   #FRK_Route_DeclarationCell := FALSE;
   IF NOT "FRK_PathOwned"(OwnerPath := #Module.Status.Name, TargetPath := #Request.TargetPath) THEN
       RETURN;
   END_IF;
   IF #Request.TargetPath = STRING_TO_WSTRING(#Module.Status.Name) THEN
       FOR #Index := 1 TO 16 DO
           #Module.ManConditions[#Index].Used := FALSE;
       END_FOR;
       "FRK_ManualApply"(Core := #Module.Core,
                         Status := #Module.Status,
                         Request := #Request,
                         Commands := #Module.Catalog,
                         Count := #Module.CatalogCount,
                         Conditions := #Module.ManConditions,
                         Report := #Report,
                         Execute := #Module.Execute,
                         Command := #Module.Command,
                         ManualOwned := #Module.ManualOwned);
       #FRK_Route_DeclarationCell := TRUE;
       RETURN;
   END_IF;
   #RouteMatched := "FRK_Route_DeclarationCylinder"(Module := #Module.Clamp, Hal := #Hal.Clamp, Request := #Request, Report := #Report);
   #FRK_Route_DeclarationCell := #FRK_Route_DeclarationCell OR #RouteMatched;
   #RouteMatched := "FRK_Route_DeclarationCylinder"(Module := #Module.Gate, Hal := #Hal.Gate, Request := #Request, Report := #Report);
   #FRK_Route_DeclarationCell := #FRK_Route_DeclarationCell OR #RouteMatched;
END_FUNCTION

FUNCTION "FRK_Route_DeclarationCylinder" : Bool   // FC130, SCL
{ S7_Optimized_Access := 'TRUE' }
VERSION : 0.1
// stored: AutoNumber true, IsIECCheckEnabled false, SetENOAutomatically false, UDAEnableTagReadback false
   VAR_INPUT
      Request : "ST_HmiRequest";
   END_VAR
   VAR_IN_OUT
      Module : "FB_DeclarationCylinder";
      Hal : "ST_DeclarationLeafHal";
      Report : "ST_ReleaseReport";
   END_VAR
   VAR_TEMP
      RouteMatched : Bool;
      Index : Int;
   END_VAR
BEGIN

   #FRK_Route_DeclarationCylinder := FALSE;
   IF NOT "FRK_PathOwned"(OwnerPath := #Module.Status.Name, TargetPath := #Request.TargetPath) THEN
       RETURN;
   END_IF;
   IF #Request.TargetPath = STRING_TO_WSTRING(#Module.Status.Name) THEN
       FOR #Index := 1 TO 16 DO
           #Module.ManConditions[#Index].Used := FALSE;
       END_FOR;
       // ---- AUTHORED: OnManRelease
       "FRK_ManualCondition"(Conditions := #Module.ManConditions,
                             Slot := 1,
                             Value := 2,
                             Ok := #Hal.Permit,
                             Diag := #Hal.Diag,
                             Bypassable := FALSE);
       "FRK_ManualCondition"(Conditions := #Module.ManConditions,
                             Slot := 2,
                             Value := 2,
                             Ok := #Hal.Sample = 0,
                             Diag := #Hal.LaterDiag,
                             Bypassable := FALSE);
       // ---- GENERATED: manual release end
       "FRK_ManualApply"(Core := #Module.Core,
                         Status := #Module.Status,
                         Request := #Request,
                         Commands := #Module.Catalog,
                         Count := #Module.CatalogCount,
                         Conditions := #Module.ManConditions,
                         Report := #Report,
                         Execute := #Module.Execute,
                         Command := #Module.Command,
                         ManualOwned := #Module.ManualOwned);
       #FRK_Route_DeclarationCylinder := TRUE;
       RETURN;
   END_IF;
END_FUNCTION

FUNCTION "FRK_Route_DeclarationUnit" : Bool   // FC163, SCL
{ S7_Optimized_Access := 'TRUE' }
VERSION : 0.1
// stored: AutoNumber true, IsIECCheckEnabled false, SetENOAutomatically false, UDAEnableTagReadback false
   VAR_INPUT
      Request : "ST_HmiRequest";
   END_VAR
   VAR_IN_OUT
      Module : "FB_DeclarationUnit";
      Hal : "ST_DeclarationUnitHal";
      Report : "ST_ReleaseReport";
   END_VAR
   VAR_TEMP
      RouteMatched : Bool;
      Index : Int;
   END_VAR
BEGIN

   #FRK_Route_DeclarationUnit := FALSE;
   IF NOT "FRK_PathOwned"(OwnerPath := #Module.Status.Name, TargetPath := #Request.TargetPath) THEN
       RETURN;
   END_IF;
   "FRK_Release_DeclarationUnit"(Unit := #Module.Unit,
                                 Hal := #Hal);
   "FRK_ManualCommon"(Core := #Module.Core,
                      Unit := #Module.Unit,
                      Status := #Module.Status,
                      Report := #Report);
   IF #Request.TargetPath = STRING_TO_WSTRING(#Module.Status.Name) THEN
       "FRK_ReleaseReason"(Report := #Report,
                           Description := WSTRING#'std.error.unsupportedHmiRequest',
                           Reason := 2008,
                           Path := STRING_TO_WSTRING(#Module.Status.Name),
                           Kind := 4);
       #FRK_Route_DeclarationUnit := TRUE;
       RETURN;
   END_IF;
   #RouteMatched := "FRK_Route_DeclarationCell"(Module := #Module.Cell, Hal := #Hal.Cell, Request := #Request, Report := #Report);
   #FRK_Route_DeclarationUnit := #FRK_Route_DeclarationUnit OR #RouteMatched;
   #RouteMatched := "FRK_Route_SatelliteUnit"(Module := #Module.Satellite, Hal := #Hal.Satellite, Request := #Request, Report := #Report);
   #FRK_Route_DeclarationUnit := #FRK_Route_DeclarationUnit OR #RouteMatched;
END_FUNCTION

FUNCTION "FRK_Route_InnerUnit" : Bool   // FC147, SCL
{ S7_Optimized_Access := 'TRUE' }
VERSION : 0.1
// stored: AutoNumber true, IsIECCheckEnabled false, SetENOAutomatically false, UDAEnableTagReadback false
   VAR_INPUT
      Request : "ST_HmiRequest";
   END_VAR
   VAR_IN_OUT
      Module : "FB_InnerUnit";
      Hal : "ST_InnerUnitHal";
      Report : "ST_ReleaseReport";
   END_VAR
   VAR_TEMP
      RouteMatched : Bool;
      Index : Int;
   END_VAR
BEGIN

   #FRK_Route_InnerUnit := FALSE;
   IF NOT "FRK_PathOwned"(OwnerPath := #Module.Status.Name, TargetPath := #Request.TargetPath) THEN
       RETURN;
   END_IF;
   "FRK_Release_InnerUnit"(Unit := #Module.Unit,
                           Hal := #Hal);
   "FRK_ManualCommon"(Core := #Module.Core,
                      Unit := #Module.Unit,
                      Status := #Module.Status,
                      Report := #Report);
   IF #Request.TargetPath = STRING_TO_WSTRING(#Module.Status.Name) THEN
       "FRK_ReleaseReason"(Report := #Report,
                           Description := WSTRING#'std.error.unsupportedHmiRequest',
                           Reason := 2008,
                           Path := STRING_TO_WSTRING(#Module.Status.Name),
                           Kind := 4);
       #FRK_Route_InnerUnit := TRUE;
       RETURN;
   END_IF;
   #RouteMatched := "FRK_Route_DeclarationCell"(Module := #Module.Cell, Hal := #Hal.Cell, Request := #Request, Report := #Report);
   #FRK_Route_InnerUnit := #FRK_Route_InnerUnit OR #RouteMatched;
END_FUNCTION

FUNCTION "FRK_Route_SatelliteUnit" : Bool   // FC155, SCL
{ S7_Optimized_Access := 'TRUE' }
VERSION : 0.1
// stored: AutoNumber true, IsIECCheckEnabled false, SetENOAutomatically false, UDAEnableTagReadback false
   VAR_INPUT
      Request : "ST_HmiRequest";
   END_VAR
   VAR_IN_OUT
      Module : "FB_SatelliteUnit";
      Hal : "ST_SatelliteUnitHal";
      Report : "ST_ReleaseReport";
   END_VAR
   VAR_TEMP
      RouteMatched : Bool;
      Index : Int;
   END_VAR
BEGIN

   #FRK_Route_SatelliteUnit := FALSE;
   IF NOT "FRK_PathOwned"(OwnerPath := #Module.Status.Name, TargetPath := #Request.TargetPath) THEN
       RETURN;
   END_IF;
   "FRK_Release_SatelliteUnit"(Unit := #Module.Unit,
                               Hal := #Hal);
   "FRK_ManualCommon"(Core := #Module.Core,
                      Unit := #Module.Unit,
                      Status := #Module.Status,
                      Report := #Report);
   IF #Request.TargetPath = STRING_TO_WSTRING(#Module.Status.Name) THEN
       "FRK_ReleaseReason"(Report := #Report,
                           Description := WSTRING#'std.error.unsupportedHmiRequest',
                           Reason := 2008,
                           Path := STRING_TO_WSTRING(#Module.Status.Name),
                           Kind := 4);
       #FRK_Route_SatelliteUnit := TRUE;
       RETURN;
   END_IF;
   #RouteMatched := "FRK_Route_DeclarationCell"(Module := #Module.Cell, Hal := #Hal.Cell, Request := #Request, Report := #Report);
   #FRK_Route_SatelliteUnit := #FRK_Route_SatelliteUnit OR #RouteMatched;
   #RouteMatched := "FRK_Route_InnerUnit"(Module := #Module.Inner, Hal := #Hal.Inner, Request := #Request, Report := #Report);
   #FRK_Route_SatelliteUnit := #FRK_Route_SatelliteUnit OR #RouteMatched;
END_FUNCTION

FUNCTION "FRK_SetBoot" : Void   // FC125, SCL
{ S7_Optimized_Access := 'TRUE' }
VERSION : 0.1
// stored: AutoNumber true, IsIECCheckEnabled false, SetENOAutomatically false, UDAEnableTagReadback false
   VAR_INPUT
      Startup : Bool;
   END_VAR
   VAR_TEMP
      RootIndex : Int;
      Slot : Int;
   END_VAR
BEGIN

   IF NOT #Startup THEN
       RETURN;
   END_IF;
   IF "FRK_SetStore".SchemaVersion <> 1 THEN
       FOR #RootIndex := 1 TO 2 DO
           IF "FRK_SetStore".SchemaVersion <> 0 THEN
               "FRK_ConfigLoss"(RootIndex := #RootIndex,
                                Scope := "FRK_SetStore".Sets[#RootIndex, 1].Info.RootIdentity);
           END_IF;
           FOR #Slot := 1 TO 4 DO
               "FRK_SetStore".Sets[#RootIndex, #Slot].Info.Used := FALSE;
           END_FOR;
       END_FOR;
       "FRK_SetStore".SchemaVersion := 1;
   END_IF;
END_FUNCTION

FUNCTION "FRK_SetCheck" : Int   // FC115, SCL
{ S7_Optimized_Access := 'TRUE' }
VERSION : 0.1
// stored: AutoNumber true, IsIECCheckEnabled false, SetENOAutomatically false, UDAEnableTagReadback false
   VAR_INPUT
      RootIndex : Int;
      Scope : String;
      Access : "FRK_Access";
      Ready : Bool;
      WriteAccess : Bool;
   END_VAR
   VAR_TEMP
      Index : Int;
      Ok : Bool;
   END_VAR
BEGIN

   #FRK_SetCheck := 0;
   "FRK_SetRuntime".Work[#RootIndex].RejectScope := #Scope;
   "FRK_SetRuntime".Work[#RootIndex].RejectKey := "FRK_ConfigScratch".Entry.WriteKey;
   #Index := "FRK_SetRecord"(RootIndex := #RootIndex, Scope := #Scope, WriteKey := "FRK_ConfigScratch".Entry.WriteKey);
   IF #Index = 0 THEN
       RETURN;
   END_IF;
   IF #Access.CurrentLevel < MAX(IN1 := #Access.Policy.Required[0], IN2 := "FRK_ConfigScratch".MinRead) THEN
       RETURN;
   END_IF;
   IF #WriteAccess THEN
       IF #Access.CurrentLevel < MAX(IN1 := #Access.Policy.Required[1], IN2 := "FRK_ConfigScratch".MinWrite) THEN
           RETURN;
       END_IF;
       IF "FRK_ConfigScratch".Entry.RequiresReady AND NOT #Ready THEN
           RETURN;
       END_IF;
   END_IF;
   IF "FRK_SetRuntime".Work[#RootIndex].Payload.Records[#Index].Revision <> "FRK_ConfigScratch".Entry.WriteRevision
       OR "FRK_SetRuntime".Work[#RootIndex].Payload.Records[#Index].Kind <> "FRK_ConfigScratch".Entry.ConfigKind
       OR "FRK_SetRuntime".Work[#RootIndex].Payload.Records[#Index].ValueType <> "FRK_ConfigScratch".Entry.ValueType THEN
       RETURN;
   END_IF;
   #Ok := "FRK_ConfigDecode"(Text := STRING_TO_WSTRING("FRK_SetRuntime".Work[#RootIndex].Payload.Records[#Index].ValueText), Storage := "FRK_ConfigScratch".Storage,
                             Minimum := "FRK_ConfigScratch".Minimum, Maximum := "FRK_ConfigScratch".Maximum, MaxLength := "FRK_ConfigScratch".MaxLength, Value := "FRK_ConfigScratch".Value);
   IF NOT #Ok THEN
       RETURN;
   END_IF;
   // Existing keyed slots are reserved before commit: commit cannot allocate.
   IF #WriteAccess AND "FRK_ConfigFind"(Scope := #Scope, Key := "FRK_ConfigScratch".Entry.WriteKey, ModelCode := "FRK_SetRuntime".Work[#RootIndex].Payload.Info.ModelCode) = 0 THEN
       RETURN;
   END_IF;
   "FRK_SetRuntime".Work[#RootIndex].Seen[#Index] := TRUE;
   "FRK_SetRuntime".Work[#RootIndex].Matched := "FRK_SetRuntime".Work[#RootIndex].Matched + 1;
   #FRK_SetCheck := #Index;
END_FUNCTION

FUNCTION "FRK_SetFind" : Int   // FC112, SCL
{ S7_Optimized_Access := 'TRUE' }
VERSION : 0.1
// Deployment-sized keyed set storage; validation belongs to the typed walk.
// stored: AutoNumber true, IsIECCheckEnabled false, SetENOAutomatically false, UDAEnableTagReadback false
   VAR_INPUT
      RootIndex : Int;
      SetName : String;
   END_VAR
   VAR_TEMP
      Index : Int;
   END_VAR
BEGIN

   #FRK_SetFind := 0;
   FOR #Index := 1 TO 4 DO
       IF "FRK_SetStore".Sets[#RootIndex, #Index].Info.Used AND "FRK_SetStore".Sets[#RootIndex, #Index].Info.SetName = #SetName THEN
           #FRK_SetFind := #Index;
           RETURN;
       END_IF;
   END_FOR;
END_FUNCTION

FUNCTION "FRK_SetIdentity" : Void   // FC2, SCL
{ S7_Optimized_Access := 'TRUE' }
VERSION : 0.1
// Generated registry services v0.1; compact rows contain no operator strings.
// stored: AutoNumber true, IsIECCheckEnabled false, SetENOAutomatically false, UDAEnableTagReadback false
   VAR_INPUT
      InstancePath : WString;
      ModuleType : DInt;
      TypeId : DInt;
      Capabilities : DWord;
      ParentIndex : DInt;
      TypeKey : String;
   END_VAR
   VAR_IN_OUT
      Core : "FRK_Core";
      Status : "ST_ModuleStatus";
   END_VAR
   VAR_TEMP
      Identity : String[254];
      QuotePos : Int;
      RowIndex : DInt;
   END_VAR
BEGIN

   #Core.Named := TRUE;
   #Core.RegIndex := 0;
   IF "FRK_Registry".Fault OR "FRK_Registry".Count < 0 OR "FRK_Registry".Count > 32
       OR #ParentIndex < 0 OR #ParentIndex > "FRK_Registry".Count OR #ParentIndex > 32 THEN
       "FRK_Registry".Fault := TRUE;
       RETURN;
   END_IF;
   IF #ParentIndex > 0 THEN
       IF NOT "FRK_Registry".Rows[#ParentIndex].Valid THEN
           "FRK_Registry".Fault := TRUE;
           RETURN;
       END_IF;
   END_IF;
   IF LEN(#InstancePath) > 254 THEN
       "FRK_Registry".Fault := TRUE;
       RETURN;
   END_IF;
   #Identity := WSTRING_TO_STRING(#InstancePath);
   #QuotePos := FIND(IN1 := #Identity, IN2 := '"');
   WHILE #QuotePos > 0 DO
       #Identity := DELETE(IN := #Identity, L := 1, P := #QuotePos);
       #QuotePos := FIND(IN1 := #Identity, IN2 := '"');
   END_WHILE;
   IF LEN(#Identity) > 80 OR LEN(#Identity) = 0 OR "FRK_Registry".Count >= 32 THEN
       "FRK_Registry".Fault := TRUE;
       RETURN;
   END_IF;
   "FRK_Registry".Count := "FRK_Registry".Count + 1;
   #RowIndex := "FRK_Registry".Count;
   #Core.RegIndex := #RowIndex;
   #Core.ParentIndex := #ParentIndex;
   #Core.ModuleType := #ModuleType;
   #Status.Name := #Identity;
   #Status.TypeKey := #TypeKey;
   #Status.ModuleType := #ModuleType;
   #Status.TileEnable := TRUE;
   "FRK_Registry".Rows[#RowIndex].Valid := TRUE;
   "FRK_Registry".Rows[#RowIndex].Parent := #ParentIndex;
   "FRK_Registry".Rows[#RowIndex].ModuleType := #ModuleType;
   "FRK_Registry".Rows[#RowIndex].TypeId := #TypeId;
   "FRK_Registry".Rows[#RowIndex].Capabilities := #Capabilities;
END_FUNCTION

FUNCTION "FRK_SetImport" : Bool   // FC120, SCL
{ S7_Optimized_Access := 'TRUE' }
VERSION : 0.1
// stored: AutoNumber true, IsIECCheckEnabled false, SetENOAutomatically false, UDAEnableTagReadback false
   VAR_INPUT
      RootIndex : Int;
      Request : "ST_HmiRequest";
   END_VAR
   VAR_TEMP
      Ok : Bool;
      Index : Int;
   END_VAR
BEGIN

   #FRK_SetImport := FALSE;
   IF #Request.IntValue <> 0 AND #Request.IntValue <> 1 THEN
       RETURN;
   END_IF;
   IF #Request.NameValue <> '' OR #Request.TargetPath <> WSTRING#'' OR #Request.DurationMs <> 0 THEN
       RETURN;
   END_IF;
   #Ok := "FRK_JsonPut"(Text := #Request.TextValue, Line := "FRK_SetRuntime".Work[#RootIndex].Piece);
   IF NOT #Ok THEN
       RETURN;
   END_IF;
   IF #Request.IntValue = 1 THEN
       #FRK_SetImport := NOT #Request.BoolValue;
       RETURN;
   END_IF;
   "FRK_SetRuntime".Work[#RootIndex].Line := "FRK_SetRuntime".Work[#RootIndex].Piece;
   "FRK_SetRuntime".Work[#RootIndex].Piece := WSTRING#'';
   #Ok := "FRK_JsonParse"(Line := "FRK_SetRuntime".Work[#RootIndex].Line, Fields := "FRK_SetRuntime".Work[#RootIndex].Fields, Count := "FRK_SetRuntime".Work[#RootIndex].FieldCount);
   IF NOT #Ok THEN
       RETURN;
   END_IF;
   IF NOT "FRK_SetRuntime".Work[#RootIndex].Importing THEN
       #Ok := "FRK_JsonReadHeader"(Count := "FRK_SetRuntime".Work[#RootIndex].FieldCount,
                                   Fields := "FRK_SetRuntime".Work[#RootIndex].Fields,
                                   Data := "FRK_SetRuntime".Work[#RootIndex].Payload.Info);
       IF NOT #Ok OR #Request.BoolValue THEN
           RETURN;
       END_IF;
       "FRK_SetRuntime".Work[#RootIndex].Payload.Info.Used := TRUE;
       "FRK_SetRuntime".Work[#RootIndex].Received := 0;
       "FRK_SetRuntime".Work[#RootIndex].Importing := TRUE;
   ELSE
       #Index := "FRK_SetRuntime".Work[#RootIndex].Received + 1;
       IF #Index > 24 OR #Index > "FRK_SetRuntime".Work[#RootIndex].Payload.Info.RecordCount THEN
           RETURN;
       END_IF;
       #Ok := "FRK_JsonReadRecord"(Count := "FRK_SetRuntime".Work[#RootIndex].FieldCount,
                                   Fields := "FRK_SetRuntime".Work[#RootIndex].Fields,
                                   Data := "FRK_SetRuntime".Work[#RootIndex].Payload.Records[#Index]);
       IF NOT #Ok THEN
           RETURN;
       END_IF;
       "FRK_SetRuntime".Work[#RootIndex].Received := #Index;
   END_IF;
   IF #Request.BoolValue THEN
       "FRK_SetRuntime".Work[#RootIndex].Importing := FALSE;
       IF "FRK_SetRuntime".Work[#RootIndex].Received <> "FRK_SetRuntime".Work[#RootIndex].Payload.Info.RecordCount THEN
           RETURN;
       END_IF;
   END_IF;
   #FRK_SetImport := TRUE;
END_FUNCTION

FUNCTION "FRK_SetRecord" : Int   // FC114, SCL
{ S7_Optimized_Access := 'TRUE' }
VERSION : 0.1
// stored: AutoNumber true, IsIECCheckEnabled false, SetENOAutomatically false, UDAEnableTagReadback false
   VAR_INPUT
      RootIndex : Int;
      Scope : String;
      WriteKey : String;
   END_VAR
   VAR_TEMP
      Index : Int;
   END_VAR
BEGIN

   #FRK_SetRecord := 0;
   FOR #Index := 1 TO "FRK_SetRuntime".Work[#RootIndex].Payload.Info.RecordCount DO
       IF "FRK_SetRuntime".Work[#RootIndex].Payload.Records[#Index].Scope = #Scope AND "FRK_SetRuntime".Work[#RootIndex].Payload.Records[#Index].WriteKey = #WriteKey THEN
           #FRK_SetRecord := #Index;
           RETURN;
       END_IF;
   END_FOR;
END_FUNCTION

FUNCTION "FRK_SetResult" : Void   // FC124, SCL
{ S7_Optimized_Access := 'TRUE' }
VERSION : 0.1
// stored: AutoNumber true, IsIECCheckEnabled false, SetENOAutomatically false, UDAEnableTagReadback false
   VAR_INPUT
      Request : "ST_HmiRequest";
      Response : "ST_HmiResponse";
      Scope : String;
      RootIndex : Int;
   END_VAR
   VAR_IN_OUT
      Persist : "ST_ConfigPersistStatus";
      AlarmLog : "FRK_AlarmLog";
   END_VAR
   VAR_TEMP
      Diag : "ST_Diagnostic";
      Slot : Int;
      Ok : Bool;
   END_VAR
BEGIN

   IF #Request.Kind <> 29 THEN
       RETURN;
   END_IF;
   IF NOT #Response.Accepted THEN
       #Persist.LastRejectScope := "FRK_SetRuntime".Work[#RootIndex].RejectScope;
       #Persist.LastRejectKey := "FRK_SetRuntime".Work[#RootIndex].RejectKey;
   END_IF;
   #Diag := "FRK_UnitScratch".EmptyDiagnostic;
   #Diag.SourcePath := STRING_TO_WSTRING(#Scope);
   IF #Response.Accepted THEN
       #Diag.ReasonCode := 2043;
       #Diag.Description := WSTRING#'std.event.configSetApplied';
   ELSE
       #Diag.ReasonCode := 2042;
       #Diag.Description := WSTRING#'std.error.configSetRejected';
       #Diag.SourcePath := STRING_TO_WSTRING(#Persist.LastRejectScope);
   END_IF;
   #Slot := "FRK_AlarmRaise"(AlarmLog := #AlarmLog, Diag := #Diag, ResetClass := 0);
   IF #Slot > 0 THEN
       #Ok := "FRK_AlarmGone"(AlarmLog := #AlarmLog, Slot := #Slot);
   END_IF;
END_FUNCTION

FUNCTION "FRK_SetShape" : Bool   // FC119, SCL
{ S7_Optimized_Access := 'TRUE' }
VERSION : 0.1
// stored: AutoNumber true, IsIECCheckEnabled false, SetENOAutomatically false, UDAEnableTagReadback false
   VAR_INPUT
      RootIndex : Int;
      RootIdentity : String;
   END_VAR
   VAR_TEMP
      Index : Int;
      Other : Int;
      ModelIndex : Int;
      KnownModel : Bool;
   END_VAR
BEGIN

   #FRK_SetShape := FALSE;
   IF NOT "FRK_SetRuntime".Work[#RootIndex].Payload.Info.Used OR "FRK_SetRuntime".Work[#RootIndex].Payload.Info.RootIdentity <> #RootIdentity
       OR "FRK_SetRuntime".Work[#RootIndex].Payload.Info.SetSchema <> 1 OR "FRK_SetRuntime".Work[#RootIndex].Payload.Info.ConfigRev = 0
       OR LEN("FRK_SetRuntime".Work[#RootIndex].Payload.Info.SetName) = 0
       OR "FRK_SetRuntime".Work[#RootIndex].Payload.Info.RecordCount < 1 OR "FRK_SetRuntime".Work[#RootIndex].Payload.Info.RecordCount > 24 THEN
       RETURN;
   END_IF;
   IF "FRK_SetRuntime".Work[#RootIndex].Payload.Info.Kind = 0 THEN
       #KnownModel := FALSE;
       FOR #ModelIndex := 1 TO 2 DO
           IF "FRK_SetRuntime".Work[#RootIndex].Payload.Info.ModelCode = "FRK_ConfigModelCode"(RootIndex := #RootIndex, ModelIndex := INT_TO_UDINT(#ModelIndex)) THEN
               #KnownModel := TRUE;
           END_IF;
       END_FOR;
       IF NOT #KnownModel THEN
           RETURN;
       END_IF;
   ELSIF "FRK_SetRuntime".Work[#RootIndex].Payload.Info.Kind <> 1 OR "FRK_SetRuntime".Work[#RootIndex].Payload.Info.ModelCode <> '' THEN
       RETURN;
   END_IF;
   FOR #Index := 1 TO "FRK_SetRuntime".Work[#RootIndex].Payload.Info.RecordCount DO
       "FRK_SetRuntime".Work[#RootIndex].RejectScope := "FRK_SetRuntime".Work[#RootIndex].Payload.Records[#Index].Scope;
       "FRK_SetRuntime".Work[#RootIndex].RejectKey := "FRK_SetRuntime".Work[#RootIndex].Payload.Records[#Index].WriteKey;
       IF "FRK_SetRuntime".Work[#RootIndex].Payload.Records[#Index].Kind <> "FRK_SetRuntime".Work[#RootIndex].Payload.Info.Kind THEN
           RETURN;
       END_IF;
       FOR #Other := 1 TO #Index - 1 DO
           IF "FRK_SetRuntime".Work[#RootIndex].Payload.Records[#Other].Scope = "FRK_SetRuntime".Work[#RootIndex].Payload.Records[#Index].Scope
               AND "FRK_SetRuntime".Work[#RootIndex].Payload.Records[#Other].WriteKey = "FRK_SetRuntime".Work[#RootIndex].Payload.Records[#Index].WriteKey THEN
               RETURN;
           END_IF;
       END_FOR;
   END_FOR;
   #FRK_SetShape := TRUE;
END_FUNCTION

FUNCTION "FRK_SetSlot" : Int   // FC113, SCL
{ S7_Optimized_Access := 'TRUE' }
VERSION : 0.1
// stored: AutoNumber true, IsIECCheckEnabled false, SetENOAutomatically false, UDAEnableTagReadback false
   VAR_INPUT
      RootIndex : Int;
      SetName : String;
   END_VAR
   VAR_TEMP
      Index : Int;
   END_VAR
BEGIN

   #FRK_SetSlot := "FRK_SetFind"(RootIndex := #RootIndex, SetName := #SetName);
   IF #FRK_SetSlot <> 0 THEN
       RETURN;
   END_IF;
   FOR #Index := 1 TO 4 DO
       IF NOT "FRK_SetStore".Sets[#RootIndex, #Index].Info.Used THEN
           #FRK_SetSlot := #Index;
           RETURN;
       END_IF;
   END_FOR;
END_FUNCTION

FUNCTION "FRK_SetValidateBegin" : Void   // FC122, SCL
{ S7_Optimized_Access := 'TRUE' }
VERSION : 0.1
// stored: AutoNumber true, IsIECCheckEnabled false, SetENOAutomatically false, UDAEnableTagReadback false
   VAR_INPUT
      RootIndex : Int;
   END_VAR
   VAR_TEMP
      Index : Int;
   END_VAR
BEGIN

   "FRK_SetRuntime".Work[#RootIndex].Matched := 0;
   FOR #Index := 1 TO 24 DO
       "FRK_SetRuntime".Work[#RootIndex].Seen[#Index] := FALSE;
   END_FOR;
END_FUNCTION

FUNCTION "FRK_SetValidateEnd" : Bool   // FC123, SCL
{ S7_Optimized_Access := 'TRUE' }
VERSION : 0.1
// stored: AutoNumber true, IsIECCheckEnabled false, SetENOAutomatically false, UDAEnableTagReadback false
   VAR_INPUT
      RootIndex : Int;
   END_VAR
   VAR_TEMP
      Index : Int;
   END_VAR
BEGIN

   #FRK_SetValidateEnd := FALSE;
   FOR #Index := 1 TO "FRK_SetRuntime".Work[#RootIndex].Payload.Info.RecordCount DO
       IF NOT "FRK_SetRuntime".Work[#RootIndex].Seen[#Index] THEN
           "FRK_SetRuntime".Work[#RootIndex].RejectScope := "FRK_SetRuntime".Work[#RootIndex].Payload.Records[#Index].Scope;
           "FRK_SetRuntime".Work[#RootIndex].RejectKey := "FRK_SetRuntime".Work[#RootIndex].Payload.Records[#Index].WriteKey;
           RETURN;
       END_IF;
   END_FOR;
   #FRK_SetValidateEnd := "FRK_SetRuntime".Work[#RootIndex].Matched = "FRK_SetRuntime".Work[#RootIndex].Payload.Info.RecordCount;
END_FUNCTION

FUNCTION "FRK_Sha256Pin" : Bool   // FC47, SCL
{ S7_Optimized_Access := 'TRUE' }
VERSION : 0.1
// Core section 7.7 prototype: private retained provider injection and independent root sessions.
//  User records are salted Core-compatible hashes, never commissioning plaintext.
// stored: AutoNumber true, IsIECCheckEnabled false, SetENOAutomatically false, UDAEnableTagReadback false
   VAR_INPUT
      Size : DInt;
   END_VAR
   VAR_IN_OUT
      Data : Array[0..47] of Byte;
      Digest : Array[0..31] of Byte;
   END_VAR
   VAR_TEMP
      BlockBytes : Array[0..63] of Byte;
      Words : Array[0..63] of DWord;
      Hash : Array[0..7] of DWord;
      Index : DInt;
      "A" : DWord;
      "B" : DWord;
      C : DWord;
      D : DWord;
      "E" : DWord;
      F : DWord;
      G : DWord;
      H : DWord;
      S0 : DWord;
      S1 : DWord;
      T1 : DWord;
      T2 : DWord;
      K : Array[0..63] of DWord;
   END_VAR
BEGIN

   #FRK_Sha256Pin := FALSE;
   #K[0] := DWORD#16#428A2F98;
   #K[1] := DWORD#16#71374491;
   #K[2] := DWORD#16#B5C0FBCF;
   #K[3] := DWORD#16#E9B5DBA5;
   #K[4] := DWORD#16#3956C25B;
   #K[5] := DWORD#16#59F111F1;
   #K[6] := DWORD#16#923F82A4;
   #K[7] := DWORD#16#AB1C5ED5;
   #K[8] := DWORD#16#D807AA98;
   #K[9] := DWORD#16#12835B01;
   #K[10] := DWORD#16#243185BE;
   #K[11] := DWORD#16#550C7DC3;
   #K[12] := DWORD#16#72BE5D74;
   #K[13] := DWORD#16#80DEB1FE;
   #K[14] := DWORD#16#9BDC06A7;
   #K[15] := DWORD#16#C19BF174;
   #K[16] := DWORD#16#E49B69C1;
   #K[17] := DWORD#16#EFBE4786;
   #K[18] := DWORD#16#0FC19DC6;
   #K[19] := DWORD#16#240CA1CC;
   #K[20] := DWORD#16#2DE92C6F;
   #K[21] := DWORD#16#4A7484AA;
   #K[22] := DWORD#16#5CB0A9DC;
   #K[23] := DWORD#16#76F988DA;
   #K[24] := DWORD#16#983E5152;
   #K[25] := DWORD#16#A831C66D;
   #K[26] := DWORD#16#B00327C8;
   #K[27] := DWORD#16#BF597FC7;
   #K[28] := DWORD#16#C6E00BF3;
   #K[29] := DWORD#16#D5A79147;
   #K[30] := DWORD#16#06CA6351;
   #K[31] := DWORD#16#14292967;
   #K[32] := DWORD#16#27B70A85;
   #K[33] := DWORD#16#2E1B2138;
   #K[34] := DWORD#16#4D2C6DFC;
   #K[35] := DWORD#16#53380D13;
   #K[36] := DWORD#16#650A7354;
   #K[37] := DWORD#16#766A0ABB;
   #K[38] := DWORD#16#81C2C92E;
   #K[39] := DWORD#16#92722C85;
   #K[40] := DWORD#16#A2BFE8A1;
   #K[41] := DWORD#16#A81A664B;
   #K[42] := DWORD#16#C24B8B70;
   #K[43] := DWORD#16#C76C51A3;
   #K[44] := DWORD#16#D192E819;
   #K[45] := DWORD#16#D6990624;
   #K[46] := DWORD#16#F40E3585;
   #K[47] := DWORD#16#106AA070;
   #K[48] := DWORD#16#19A4C116;
   #K[49] := DWORD#16#1E376C08;
   #K[50] := DWORD#16#2748774C;
   #K[51] := DWORD#16#34B0BCB5;
   #K[52] := DWORD#16#391C0CB3;
   #K[53] := DWORD#16#4ED8AA4A;
   #K[54] := DWORD#16#5B9CCA4F;
   #K[55] := DWORD#16#682E6FF3;
   #K[56] := DWORD#16#748F82EE;
   #K[57] := DWORD#16#78A5636F;
   #K[58] := DWORD#16#84C87814;
   #K[59] := DWORD#16#8CC70208;
   #K[60] := DWORD#16#90BEFFFA;
   #K[61] := DWORD#16#A4506CEB;
   #K[62] := DWORD#16#BEF9A3F7;
   #K[63] := DWORD#16#C67178F2;
   FOR #Index := 0 TO 31 DO
       #Digest[#Index] := 0;
   END_FOR;
   IF #Size < 0 OR #Size > 48 THEN
       RETURN;
   END_IF;
   // Authentication messages fit exactly one SHA-256 block.
   FOR #Index := 0 TO 63 DO
       #BlockBytes[#Index] := 0;
   END_FOR;
   FOR #Index := 0 TO #Size - 1 DO
       #BlockBytes[#Index] := #Data[#Index];
   END_FOR;
   #BlockBytes[#Size] := BYTE#16#80;
   #BlockBytes[62] := DWORD_TO_BYTE(SHR(IN := DINT_TO_DWORD(#Size * 8), N := 8));
   #BlockBytes[63] := DINT_TO_BYTE(#Size * 8);
   #Hash[0] := DWORD#16#6A09E667;
   #Hash[1] := DWORD#16#BB67AE85;
   #Hash[2] := DWORD#16#3C6EF372;
   #Hash[3] := DWORD#16#A54FF53A;
   #Hash[4] := DWORD#16#510E527F;
   #Hash[5] := DWORD#16#9B05688C;
   #Hash[6] := DWORD#16#1F83D9AB;
   #Hash[7] := DWORD#16#5BE0CD19;
   FOR #Index := 0 TO 15 DO
       #Words[#Index] := SHL(IN := BYTE_TO_DWORD(#BlockBytes[4 * #Index]), N := 24)
       OR SHL(IN := BYTE_TO_DWORD(#BlockBytes[4 * #Index + 1]), N := 16)
       OR SHL(IN := BYTE_TO_DWORD(#BlockBytes[4 * #Index + 2]), N := 8)
       OR BYTE_TO_DWORD(#BlockBytes[4 * #Index + 3]);
   END_FOR;
   FOR #Index := 16 TO 63 DO
       #S0 := ROR(IN := #Words[#Index - 15], N := 7) XOR ROR(IN := #Words[#Index - 15], N := 18) XOR SHR(IN := #Words[#Index - 15], N := 3);
       #S1 := ROR(IN := #Words[#Index - 2], N := 17) XOR ROR(IN := #Words[#Index - 2], N := 19) XOR SHR(IN := #Words[#Index - 2], N := 10);
       #Words[#Index] := UDINT_TO_DWORD(ULINT_TO_UDINT(UDINT_TO_ULINT(DWORD_TO_UDINT(#Words[#Index - 16])) + UDINT_TO_ULINT(DWORD_TO_UDINT(#S0)) + UDINT_TO_ULINT(DWORD_TO_UDINT(#Words[#Index - 7])) + UDINT_TO_ULINT(DWORD_TO_UDINT(#S1))));
   END_FOR;
   #A := #Hash[0];
   #B := #Hash[1];
   #C := #Hash[2];
   #D := #Hash[3];
   #E := #Hash[4];
   #F := #Hash[5];
   #G := #Hash[6];
   #H := #Hash[7];
   FOR #Index := 0 TO 63 DO
       #S1 := ROR(IN := #E, N := 6) XOR ROR(IN := #E, N := 11) XOR ROR(IN := #E, N := 25);
       #T1 := UDINT_TO_DWORD(ULINT_TO_UDINT(UDINT_TO_ULINT(DWORD_TO_UDINT(#H)) + UDINT_TO_ULINT(DWORD_TO_UDINT(#S1)) + UDINT_TO_ULINT(DWORD_TO_UDINT((#E AND #F) XOR ((NOT #E) AND #G))) + UDINT_TO_ULINT(DWORD_TO_UDINT(#K[#Index])) + UDINT_TO_ULINT(DWORD_TO_UDINT(#Words[#Index]))));
       #S0 := ROR(IN := #A, N := 2) XOR ROR(IN := #A, N := 13) XOR ROR(IN := #A, N := 22);
       #T2 := UDINT_TO_DWORD(ULINT_TO_UDINT(UDINT_TO_ULINT(DWORD_TO_UDINT(#S0)) + UDINT_TO_ULINT(DWORD_TO_UDINT((#A AND #B) XOR (#A AND #C) XOR (#B AND #C)))));
       #H := #G;
       #G := #F;
       #F := #E;
       #E := UDINT_TO_DWORD(ULINT_TO_UDINT(UDINT_TO_ULINT(DWORD_TO_UDINT(#D)) + UDINT_TO_ULINT(DWORD_TO_UDINT(#T1))));
       #D := #C;
       #C := #B;
       #B := #A;
       #A := UDINT_TO_DWORD(ULINT_TO_UDINT(UDINT_TO_ULINT(DWORD_TO_UDINT(#T1)) + UDINT_TO_ULINT(DWORD_TO_UDINT(#T2))));
   END_FOR;
   #Words[0] := #A;
   #Words[1] := #B;
   #Words[2] := #C;
   #Words[3] := #D;
   #Words[4] := #E;
   #Words[5] := #F;
   #Words[6] := #G;
   #Words[7] := #H;
   FOR #Index := 0 TO 7 DO
       #Hash[#Index] := UDINT_TO_DWORD(ULINT_TO_UDINT(UDINT_TO_ULINT(DWORD_TO_UDINT(#Hash[#Index])) + UDINT_TO_ULINT(DWORD_TO_UDINT(#Words[#Index]))));
       #Digest[4 * #Index] := DWORD_TO_BYTE(SHR(IN := #Hash[#Index], N := 24));
       #Digest[4 * #Index + 1] := DWORD_TO_BYTE(SHR(IN := #Hash[#Index], N := 16));
       #Digest[4 * #Index + 2] := DWORD_TO_BYTE(SHR(IN := #Hash[#Index], N := 8));
       #Digest[4 * #Index + 3] := DWORD_TO_BYTE(#Hash[#Index]);
   END_FOR;
   FOR #Index := 0 TO 63 DO
       #BlockBytes[#Index] := 0;
       #Words[#Index] := 0;
   END_FOR;
   #FRK_Sha256Pin := TRUE;
END_FUNCTION

FUNCTION "FRK_Start" : Void   // FC15, SCL
{ S7_Optimized_Access := 'TRUE' }
VERSION : 0.1
// stored: AutoNumber true, IsIECCheckEnabled false, SetENOAutomatically false, UDAEnableTagReadback false
   VAR_INPUT
      Supported : Bool;
      Timeout : Time;
      Label : String;
   END_VAR
   VAR_IN_OUT
      Core : "FRK_Core";
      Status : "ST_ModuleStatus";
   END_VAR
BEGIN

   #Core.CommandLabel := #Label;
   IF NOT #Supported THEN
       "FRK_Fault"(Core := #Core,
                   Status := #Status,
                   ReasonCode := 2008,
                   Description := WSTRING#'fraktal.command.unsupported');
   ELSIF #Timeout <= T#0ms THEN
       "FRK_Fault"(Core := #Core,
                   Status := #Status,
                   ReasonCode := 2004,
                   Description := WSTRING#'fraktal.command.timeout.invalid');
   ELSE
       #Core.TimeoutMs := DINT_TO_UDINT(TIME_TO_DINT(#Timeout));
   END_IF;
END_FUNCTION

FUNCTION "FRK_State" : Bool   // FC22, SCL
{ S7_Optimized_Access := 'TRUE' }
VERSION : 0.1
// stored: AutoNumber true, IsIECCheckEnabled false, SetENOAutomatically false, UDAEnableTagReadback false
   VAR_INPUT
      Idx : Int;
      Key : String;
      Ok : Bool;
   END_VAR
   VAR_IN_OUT
      Flags : Array[1..12] of "ST_StateFlag";
      Count : Int;
      Touched : Array[1..12] of Bool;
   END_VAR
   VAR_TEMP
      Stamp : DTL;
      ResultCode : Int;
   END_VAR
BEGIN

   #FRK_State := #Ok;
   IF #Idx < 1 OR #Idx > 12 OR LEN(#Key) = 0 OR LEN(#Key) > 120 THEN
       RETURN;
   END_IF;
   IF #Idx > #Count THEN
       #Count := #Idx;
   END_IF;
   IF #Flags[#Idx].Value <> #Ok OR #Flags[#Idx].Key <> #Key OR #Flags[#Idx].Stale THEN
       #Flags[#Idx].Since := LDT#1970-01-01-00:00:00.000000000;
       #ResultCode := RD_SYS_T(OUT => #Stamp);
       IF #ResultCode = 0 THEN
           #Flags[#Idx].Since := DTL_TO_LDT(#Stamp);
       END_IF;
   END_IF;
   #Flags[#Idx].Key := #Key;
   #Flags[#Idx].Value := #Ok;
   #Flags[#Idx].Stale := FALSE;
   #Touched[#Idx] := TRUE;
END_FUNCTION

FUNCTION "FRK_StateSweep" : Void   // FC21, SCL
{ S7_Optimized_Access := 'TRUE' }
VERSION : 0.1
// Core 3.12: derived facts; owning frame resolves freshness every scan.
// stored: AutoNumber true, IsIECCheckEnabled false, SetENOAutomatically false, UDAEnableTagReadback false
   VAR_INPUT
      Startup : Bool;
   END_VAR
   VAR_IN_OUT
      Flags : Array[1..12] of "ST_StateFlag";
      Count : Int;
      Touched : Array[1..12] of Bool;
   END_VAR
   VAR_TEMP
      Index : Int;
   END_VAR
BEGIN

   IF #Count < 0 OR #Count > 12 THEN
       #Count := 0;
   END_IF;
   FOR #Index := 1 TO #Count DO
       IF #Startup OR NOT #Touched[#Index] THEN
           #Flags[#Index].Value := FALSE;
           #Flags[#Index].Stale := TRUE;
       END_IF;
       #Touched[#Index] := FALSE;
   END_FOR;
END_FUNCTION

FUNCTION "FRK_SyncRegistry" : Void   // FC3, SCL
{ S7_Optimized_Access := 'TRUE' }
VERSION : 0.1
// stored: AutoNumber true, IsIECCheckEnabled false, SetENOAutomatically false, UDAEnableTagReadback false
   VAR_INPUT
      Index : DInt;
      Status : "ST_ModuleStatus";
   END_VAR
BEGIN

   // Nested checks precede array access; do not depend on short-circuit AND.
   IF #Index < 1 OR #Index > "FRK_Registry".Count OR #Index > 32 THEN
       "FRK_Registry".Fault := TRUE;
       RETURN;
   END_IF;
   IF NOT "FRK_Registry".Rows[#Index].Valid THEN
       "FRK_Registry".Fault := TRUE;
       RETURN;
   END_IF;
   "FRK_Registry".Rows[#Index].Exec := #Status.State;
   "FRK_Registry".Rows[#Index].ReasonCode := #Status.Diagnostic.ReasonCode;
   "FRK_Registry".Rows[#Index].Severity := #Status.Diagnostic.Severity;
END_FUNCTION

FUNCTION "FRK_UnitCascade" : Void   // FC92, SCL
{ S7_Optimized_Access := 'TRUE' }
VERSION : 0.1
// stored: AutoNumber true, IsIECCheckEnabled false, SetENOAutomatically false, UDAEnableTagReadback false
   VAR_INPUT
      ParentUnit : "FRK_Unit";
      Supported : Array[0..6] of Bool;
   END_VAR
   VAR_IN_OUT
      Core : "FRK_Core";
      Unit : "FRK_Unit";
      Status : "ST_ModuleStatus";
      Policy : Array[0..6] of "ST_ModePolicy";
      Access : "FRK_Access";
      AlarmLog : "FRK_AlarmLog";
   END_VAR
   VAR_TEMP
      Request : "ST_HmiRequest";
   END_VAR
BEGIN

   IF NOT #ParentUnit.CascadePending THEN
       RETURN;
   END_IF;
   IF #ParentUnit.CascadeKind = 6 OR #ParentUnit.CascadeKind = 9 THEN
       #Unit.FollowStart := FALSE;
       #Request.Kind := #ParentUnit.CascadeKind;
       "FRK_UnitOperation"(Core := #Core,
                           Unit := #Unit,
                           Status := #Status,
                           Policy := #Policy,
                           Access := #Access,
                           Supported := #Supported,
                           Request := #Request,
                           Response := "FRK_UnitScratch".Response,
                           Trusted := TRUE);
       RETURN;
   END_IF;
   #Request.Kind := 3;
   #Request.IntValue := #ParentUnit.CascadeMode;
   "FRK_UnitOperation"(Core := #Core,
                       Unit := #Unit,
                       Status := #Status,
                       Policy := #Policy,
                       Access := #Access,
                       Supported := #Supported,
                       Request := #Request,
                       Response := "FRK_UnitScratch".Response,
                       Trusted := TRUE);
   IF NOT "FRK_UnitScratch".Response.Accepted THEN
       #Unit.FollowStart := FALSE;
       #Request.Kind := 6;
       "FRK_UnitOperation"(Core := #Core,
                           Unit := #Unit,
                           Status := #Status,
                           Policy := #Policy,
                           Access := #Access,
                           Supported := #Supported,
                           Request := #Request,
                           Response := "FRK_UnitScratch".Response,
                           Trusted := TRUE);
       // Core names this event but has no assigned E_Reason ordinal yet.
       "FRK_AlarmMessage"(AlarmLog := #AlarmLog,
                          Reason := 2008,
                          Description := WSTRING#'std.event.childModeUnsupported',
                          SourcePath := STRING_TO_WSTRING(#Status.Name));
   ELSE
       #Unit.FollowStart := #ParentUnit.CascadeKind = 5;
   END_IF;
END_FUNCTION

FUNCTION "FRK_UnitConsume" : Void   // FC80, SCL
{ S7_Optimized_Access := 'TRUE' }
VERSION : 0.1
// stored: AutoNumber true, IsIECCheckEnabled false, SetENOAutomatically false, UDAEnableTagReadback false
   VAR_INPUT
      Supported : Array[0..6] of Bool;
   END_VAR
   VAR_IN_OUT
      Core : "FRK_Core";
      Unit : "FRK_Unit";
      Status : "ST_ModuleStatus";
      Policy : Array[0..6] of "ST_ModePolicy";
      Access : "FRK_Access";
      Response : "ST_HmiResponse";
   END_VAR
BEGIN

   IF NOT #Unit.RequestPending THEN
       RETURN;
   END_IF;
   // The generated typed ownership walk serves the static manifest after children.
   IF #Unit.Request.Kind = 23 THEN
       #Unit.Request.Secret := '';
       RETURN;
   END_IF;
   "FRK_UnitOperation"(Core := #Core,
                       Unit := #Unit,
                       Status := #Status,
                       Policy := #Policy,
                       Access := #Access,
                       Supported := #Supported,
                       Request := #Unit.Request,
                       Response := #Response,
                       Trusted := FALSE);
   #Unit.Request.Secret := '';
END_FUNCTION

FUNCTION "FRK_UnitFinish" : Void   // FC85, SCL
{ S7_Optimized_Access := 'TRUE' }
VERSION : 0.1
// stored: AutoNumber true, IsIECCheckEnabled false, SetENOAutomatically false, UDAEnableTagReadback false
   VAR_IN_OUT
      Core : "FRK_Core";
      Unit : "FRK_Unit";
      Response : "ST_HmiResponse";
      Status : "ST_ModuleStatus";
      Part : "ST_PartContext";
      AlarmLog : "FRK_AlarmLog";
      History : Array[1..16] of "ST_Diagnostic";
      Head : Int;
   END_VAR
BEGIN

   IF #Core.Exec = 3 THEN
       IF NOT #Unit.EvReset THEN
           #Unit.FaultLatched := TRUE;
       END_IF;
       IF NOT #Unit.PrevError THEN
           IF #Head < 0 OR #Head >= 16 THEN
               #Head := 0;
           END_IF;
           #Head := #Head + 1;
           #History[#Head] := #Status.Diagnostic;
           "FRK_PartAborted"(Core := #Core,
                             Unit := #Unit,
                             Status := #Status,
                             Part := #Part,
                             AlarmLog := #AlarmLog);
       END_IF;
   END_IF;
   #Unit.PrevError := #Core.Exec = 3;
   IF #Core.Exec = 2 OR #Core.Exec = 4 THEN
       #Unit.RunReq := FALSE;
   END_IF;
   IF #Unit.Clearing AND #Core.Exec = 0 THEN
       IF "FRK_DescendantsReady"(OwnerIndex := #Core.RegIndex) THEN
           #Unit.Clearing := FALSE;
       END_IF;
   END_IF;
   #Unit.AbortReq := FALSE;
   #Unit.ReleaseChildren := FALSE;
   #Unit.EvReset := FALSE;
   IF #Unit.RequestPending THEN
       #Response.AckSequence := #Unit.SeenSequence;
       #Unit.RequestPending := FALSE;
   END_IF;
END_FUNCTION

FUNCTION "FRK_UnitFollow" : Void   // FC93, SCL
{ S7_Optimized_Access := 'TRUE' }
VERSION : 0.1
// stored: AutoNumber true, IsIECCheckEnabled false, SetENOAutomatically false, UDAEnableTagReadback false
   VAR_INPUT
      Supported : Array[0..6] of Bool;
   END_VAR
   VAR_IN_OUT
      Core : "FRK_Core";
      Unit : "FRK_Unit";
      Status : "ST_ModuleStatus";
      Policy : Array[0..6] of "ST_ModePolicy";
      Access : "FRK_Access";
   END_VAR
   VAR_TEMP
      Request : "ST_HmiRequest";
   END_VAR
BEGIN

   IF #Unit.FollowStart AND NOT #Unit.ModePending AND NOT #Unit.Clearing THEN
       #Unit.FollowStart := FALSE;
       #Request.Kind := 5;
       "FRK_UnitOperation"(Core := #Core,
                           Unit := #Unit,
                           Status := #Status,
                           Policy := #Policy,
                           Access := #Access,
                           Supported := #Supported,
                           Request := #Request,
                           Response := "FRK_UnitScratch".Response,
                           Trusted := TRUE);
   END_IF;
END_FUNCTION

FUNCTION "FRK_UnitMailbox" : Void   // FC79, SCL
{ S7_Optimized_Access := 'TRUE' }
VERSION : 0.1
// stored: AutoNumber true, IsIECCheckEnabled false, SetENOAutomatically false, UDAEnableTagReadback false
   VAR_INPUT
      Supported : Array[0..6] of Bool;
   END_VAR
   VAR_IN_OUT
      Core : "FRK_Core";
      Unit : "FRK_Unit";
      Status : "ST_ModuleStatus";
      Policy : Array[0..6] of "ST_ModePolicy";
      Access : "FRK_Access";
      Request : "ST_HmiRequest";
      Response : "ST_HmiResponse";
   END_VAR
   VAR_TEMP
      SequenceBefore : UDInt;
   END_VAR
BEGIN

   #SequenceBefore := #Request.Sequence;
   IF #SequenceBefore = 0 OR #SequenceBefore = #Unit.SeenSequence THEN
       RETURN;
   END_IF;
   #Unit.Request := #Request;
   IF #Request.Sequence <> #SequenceBefore THEN
       #Unit.Request.Secret := '';
       RETURN;
   END_IF;
   #Request.Secret := '';
   #Unit.RequestUser := #Access.CurrentUser;
   #Unit.SeenSequence := #SequenceBefore;
   #Unit.RequestPending := TRUE;
END_FUNCTION

FUNCTION "FRK_UnitMode" : Void   // FC81, SCL
{ S7_Optimized_Access := 'TRUE' }
VERSION : 0.1
// stored: AutoNumber true, IsIECCheckEnabled false, SetENOAutomatically false, UDAEnableTagReadback false
   VAR_IN_OUT
      Core : "FRK_Core";
      Unit : "FRK_Unit";
   END_VAR
BEGIN

   IF #Unit.ModePending THEN
       IF #Core.Exec = 1 THEN
           #Core.EvModeExit := TRUE;
           #Core.HookResult := 0;
       ELSIF #Core.Exec = 0 AND NOT #Unit.Clearing THEN
           #Unit.Mode := #Unit.RequestedMode;
           #Unit.ModePending := FALSE;
           #Unit.ExitFirst := FALSE;
           #Core.EvModeChanged := TRUE;
       ELSE
           #Unit.RunReq := FALSE;
       END_IF;
   END_IF;
END_FUNCTION

FUNCTION "FRK_UnitModeResolve" : Void   // FC82, SCL
{ S7_Optimized_Access := 'TRUE' }
VERSION : 0.1
// stored: AutoNumber true, IsIECCheckEnabled false, SetENOAutomatically false, UDAEnableTagReadback false
   VAR_INPUT
      Policy : Array[0..6] of "ST_ModePolicy";
      Timeout : Time;
   END_VAR
   VAR_IN_OUT
      Core : "FRK_Core";
      Unit : "FRK_Unit";
      Status : "ST_ModuleStatus";
   END_VAR
BEGIN

   IF #Unit.ModePending THEN
       IF #Timeout <= T#0ms OR "FRK_Elapsed"(NewMs := "FRK_Clock".NowMs, OldMs := #Unit.ModeSince) >= DINT_TO_UDINT(TIME_TO_DINT(#Timeout)) THEN
           "FRK_Fault"(Core := #Core,
                       Status := #Status,
                       ReasonCode := 2001,
                       Description := WSTRING#'std.error.hmiRequestRejected');
           #Unit.ModePending := FALSE;
           #Unit.FollowStart := FALSE;
           #Unit.ReleaseChildren := TRUE;
           #Unit.Clearing := TRUE;
       ELSIF #Core.EvModeExit THEN
           #Unit.ExitFirst := FALSE;
           IF #Policy[#Unit.Mode].Style = 0 THEN
               #Unit.StopReq := TRUE;
           ELSIF #Core.HookResult <= 0 THEN
               #Unit.AbortReq := TRUE;
               #Unit.ReleaseChildren := TRUE;
               #Unit.Clearing := TRUE;
           END_IF;
       END_IF;
   END_IF;
END_FUNCTION

FUNCTION "FRK_UnitOperation" : Void   // FC78, SCL
{ S7_Optimized_Access := 'TRUE' }
VERSION : 0.1
// stored: AutoNumber true, IsIECCheckEnabled false, SetENOAutomatically false, UDAEnableTagReadback false
   VAR_INPUT
      Supported : Array[0..6] of Bool;
      Request : "ST_HmiRequest";
      Trusted : Bool;
   END_VAR
   VAR_IN_OUT
      Core : "FRK_Core";
      Unit : "FRK_Unit";
      Status : "ST_ModuleStatus";
      Policy : Array[0..6] of "ST_ModePolicy";
      Access : "FRK_Access";
      Response : "ST_HmiResponse";
   END_VAR
   VAR_TEMP
      Gate : DInt;
      Desired : DInt;
      Query : Bool;
      Level : DInt;
      DecisionAccepted : Bool;
   END_VAR
BEGIN

   #Response.Accepted := FALSE;
   #Response.Diagnostic := WSTRING#'';
   #Response.Report.Count := 0;
   #Response.Report.Released := TRUE;
   #Gate := -1;
   #Desired := -1;
   #Query := FALSE;
   CASE #Request.Kind OF
       5:
           #Gate := 5;
           #Desired := 0;
       6:
           #Gate := 5;
           #Desired := 1;
       3:
           #Gate := 4;
           #Desired := #Request.IntValue;
           IF #Desired = -1 THEN
               #Desired := -2;
           END_IF;
       9:
           #Gate := 7;
       10:
           #Gate := 5;
       11:
           #Gate := 2;
       24, 25:
           #Gate := 8;
       15:
           #Gate := 5;
           #Desired := 0;
           #Query := TRUE;
       16:
           #Gate := 2;
           #Query := TRUE;
       17:
           #Gate := #Request.IntValue;
           #Desired := -1;
           #Query := TRUE;
       ELSE
           #Gate := -1;
   END_CASE;
   IF #Gate <> -1 OR #Request.Kind = 17 THEN
       "FRK_UnitRelease"(Core := #Core,
                         Unit := #Unit,
                         Status := #Status,
                         Policy := #Policy,
                         Access := #Access,
                         Supported := #Supported,
                         Report := #Response.Report,
                         Gate := #Gate,
                         Desired := #Desired,
                         Trusted := #Trusted);
       IF #Query THEN
           #Response.Accepted := TRUE;
       ELSIF #Response.Report.Released THEN
           CASE #Request.Kind OF
               10:
                   #DecisionAccepted := "FRK_DecisionSubmit"(Owner := #Core.RegIndex,
                                                             OwnerPath := STRING_TO_WSTRING(#Status.Name),
                                                             Option := #Request.IntValue,
                                                             Busy := #Core.Exec = 1,
                                                             Permit := #Unit.Permit,
                                                             Report := #Response.Report);
                   #Response.Accepted := #DecisionAccepted;
               5:
                   #Unit.StopReq := FALSE;
                   #Unit.RunReq := TRUE;
                   #Response.Accepted := TRUE;
               6:
                   #Unit.StopReq := #Core.Exec = 1;
                   IF NOT #Unit.StopReq THEN
                       #Unit.RunReq := FALSE;
                   END_IF;
                   #Unit.FollowStart := FALSE;
                   #Response.Accepted := TRUE;
               3:
                   IF #Desired <> #Unit.Mode THEN
                       #Unit.ExitFirst := TRUE;
                       #Unit.ModeSince := "FRK_Clock".NowMs;
                       #Unit.RequestedMode := #Desired;
                       #Unit.ModePending := TRUE;
                       IF #Unit.Mode = 1 THEN
                           #Unit.ReleaseChildren := TRUE;
                           #Unit.Clearing := TRUE;
                       END_IF;
                   END_IF;
                   #Response.Accepted := TRUE;
               9:
                   #Unit.EvReset := TRUE;
                   #Unit.ModePending := FALSE;
                   #Unit.ExitFirst := FALSE;
                   #Unit.RunReq := FALSE;
                   #Unit.AbortReq := #Core.Exec = 1;
                   #Unit.StopReq := FALSE;
                   #Unit.FollowStart := FALSE;
                   #Unit.ReleaseChildren := TRUE;
                   #Unit.Clearing := TRUE;
                   #Unit.FaultLatched := FALSE;
                   IF #Core.Exec = 3 THEN
                       #Core.Armed := TRUE;
                   END_IF;
                   #Response.Accepted := TRUE;
               24:
                   #Level := -1;
                   IF #Request.TextValue = WSTRING#'0' THEN
                       #Level := 0;
                   ELSIF #Request.TextValue = WSTRING#'1' THEN
                       #Level := 1;
                   ELSIF #Request.TextValue = WSTRING#'2' THEN
                       #Level := 2;
                   ELSIF #Request.TextValue = WSTRING#'3' THEN
                       #Level := 3;
                   ELSIF #Request.TextValue = WSTRING#'4' THEN
                       #Level := 4;
                   END_IF;
                   IF #Request.IntValue >= 0 AND #Request.IntValue <= 11 AND #Level >= 0 THEN
                       IF #Request.IntValue <> 8 OR #Level <= #Access.CurrentLevel THEN
                           #Access.Policy.Required[#Request.IntValue] := #Level;
                           #Response.Accepted := TRUE;
                       END_IF;
                   END_IF;
               25:
                   IF #Request.DurationMs <= 604800000 THEN
                       #Access.Policy.SessionTimeout := DINT_TO_TIME(UDINT_TO_DINT(#Request.DurationMs));
                       #Response.Accepted := TRUE;
                   END_IF;
               ELSE
                   // Manual acceptance is resolved by the generated typed route.
                   #Response.Accepted := FALSE;
           END_CASE;
       END_IF;
   ELSE
       CASE #Request.Kind OF
           1:
               "FRK_AccessLogin"(Access := #Access,
                                 User := #Request.User,
                                 Secret := #Request.Secret,
                                 Sequence := #Request.Sequence);
               // Consumption is acknowledged now; correlated result is asynchronous.
               #Response.Accepted := TRUE;
           2:
               "FRK_AccessLogout"(Access := #Access);
               #Response.Accepted := TRUE;
           ELSE
               #Response.Diagnostic := WSTRING#'std.error.unsupportedHmiRequest';
       END_CASE;
   END_IF;
   IF #Response.Accepted AND NOT #Query THEN
       IF #Request.Kind = 5 OR #Request.Kind = 6 OR #Request.Kind = 3 OR #Request.Kind = 9 THEN
           #Unit.CascadePending := TRUE;
           #Unit.CascadeKind := #Request.Kind;
           #Unit.CascadeMode := #Unit.Mode;
           IF #Request.Kind = 3 THEN
               #Unit.CascadeMode := #Desired;
           END_IF;
       END_IF;
   END_IF;
   IF NOT #Response.Accepted AND #Request.Kind <> 11 THEN
       IF #Response.Diagnostic = WSTRING#'' THEN
           #Response.Diagnostic := WSTRING#'std.error.hmiRequestRejected';
       END_IF;
       IF #Response.Report.Released THEN
           "FRK_ReleaseReason"(Report := #Response.Report,
                               Description := #Response.Diagnostic,
                               Reason := 2002,
                               Path := STRING_TO_WSTRING(#Status.Name),
                               Kind := 4);
       END_IF;
   END_IF;
END_FUNCTION

FUNCTION "FRK_UnitPrepare" : Void   // FC69, SCL
{ S7_Optimized_Access := 'TRUE' }
VERSION : 0.1
// Shared Unit services v0.1: operation authority, mailbox, modes and local carrier.
// stored: AutoNumber true, IsIECCheckEnabled false, SetENOAutomatically false, UDAEnableTagReadback false
   VAR_INPUT
      Startup : Bool;
      InitialMode : DInt;
   END_VAR
   VAR_IN_OUT
      Core : "FRK_Core";
      Unit : "FRK_Unit";
      Policy : Array[0..6] of "ST_ModePolicy";
      Request : "ST_HmiRequest";
      Response : "ST_HmiResponse";
   END_VAR
   VAR_TEMP
      Index : DInt;
   END_VAR
BEGIN

   #Core.EvModeExit := FALSE;
   #Core.EvModeChanged := FALSE;
   IF NOT #Unit.Initialized THEN
       #Unit.Initialized := TRUE;
       #Unit.Permit := TRUE;
       FOR #Index := 0 TO 7 - 1 DO
           #Policy[#Index].Shield := 1;
           #Policy[#Index].Style := 1;
       END_FOR;
       #Policy[0].Style := 0;
       #Policy[2].Shield := 0;
       #Policy[1].Shield := 0;
       #Policy[3].Shield := 2;
       #Policy[4].Shield := 2;
       #Unit.Mode := #InitialMode;
   END_IF;
   IF #Startup THEN
       #Unit.EvReset := FALSE;
       #Unit.Mode := #InitialMode;
       #Unit.RunReq := FALSE;
       #Unit.AbortReq := #Core.Exec = 1;
       #Unit.StopReq := FALSE;
       #Unit.ModePending := FALSE;
       #Unit.FollowStart := FALSE;
       #Unit.CascadePending := FALSE;
       #Unit.ReleaseChildren := TRUE;
       #Unit.Clearing := TRUE;
       // Consume the restart boundary without executing a transported request.
       #Unit.SeenSequence := #Request.Sequence;
       #Unit.RequestPending := FALSE;
       #Request.Secret := '';
       #Response.Accepted := FALSE;
       #Response.Diagnostic := WSTRING#'std.error.hmiRequestRejected';
       #Response.AckSequence := #Unit.SeenSequence;
   END_IF;
   IF #Core.ReleasePending THEN
       #Unit.FollowStart := FALSE;
       // An incoming parent mode/reset operation is already queued for this scan.
       // Preserve its cascade while cancelling the old command.
       #Unit.RunReq := FALSE;
       #Unit.AbortReq := TRUE;
       #Unit.ReleaseChildren := TRUE;
       #Unit.Clearing := TRUE;
   END_IF;
END_FUNCTION

FUNCTION "FRK_UnitRelease" : Void   // FC87, SCL
{ S7_Optimized_Access := 'TRUE' }
VERSION : 0.1
// stored: AutoNumber true, IsIECCheckEnabled false, SetENOAutomatically false, UDAEnableTagReadback false
   VAR_INPUT
      Gate : DInt;
      Desired : DInt;
      Trusted : Bool;
      Core : "FRK_Core";
      Unit : "FRK_Unit";
      Status : "ST_ModuleStatus";
      Policy : Array[0..6] of "ST_ModePolicy";
      Access : "FRK_Access";
      Supported : Array[0..6] of Bool;
   END_VAR
   VAR_IN_OUT
      Report : "ST_ReleaseReport";
   END_VAR
BEGIN

   #Report.Count := 0;
   #Report.Released := TRUE;
   IF #Gate <> 5 AND #Gate <> 4
       AND #Gate <> 7 AND #Gate <> 2
       AND #Gate <> 8
       AND NOT (#Unit.ConfigEnabled AND #Gate = 1)
       AND NOT (#Unit.ConfigSetsEnabled AND #Gate = 11)
       AND NOT (#Unit.ModelEnabled AND #Gate = 3) THEN
       "FRK_ReleaseReason"(Report := #Report,
                           Description := WSTRING#'std.error.unsupportedHmiRequest',
                           Reason := 2008,
                           Path := STRING_TO_WSTRING(#Status.Name),
                           Kind := 4);
       RETURN;
   END_IF;
   IF NOT #Trusted THEN
       IF #Access.CurrentLevel < #Access.Policy.Required[#Gate] THEN
           "FRK_ReleaseReason"(Report := #Report,
                               Description := WSTRING#'std.release.insufficientAction',
                               Reason := 2002,
                               Path := STRING_TO_WSTRING(#Status.Name),
                               Kind := 1);
       END_IF;
   END_IF;
   CASE #Gate OF
       3:
           IF #Core.Exec <> 0 OR #Unit.ModePending OR #Unit.Clearing OR NOT "FRK_DescendantsReady"(OwnerIndex := #Core.RegIndex) THEN
               "FRK_ReleaseReason"(Report := #Report,
                                   Description := WSTRING#'std.error.hmiRequestRejected',
                                   Reason := 2011,
                                   Path := STRING_TO_WSTRING(#Status.Name),
                                   Kind := 4);
           END_IF;
           IF #Unit.AlarmBlocking THEN
               "FRK_ReleaseReason"(Report := #Report,
                                   Description := WSTRING#'std.release.manualReset',
                                   Reason := 0,
                                   Path := STRING_TO_WSTRING(#Status.Name),
                                   Kind := 2);
           END_IF;
           IF NOT #Unit.Permit THEN
               "FRK_ReleaseReason"(Report := #Report,
                                   Description := #Unit.PermitDiag.Description,
                                   Reason := #Unit.PermitDiag.ReasonCode,
                                   Path := #Unit.PermitDiag.SourcePath,
                                   Kind := 3);
           END_IF;
       5:
           // Desired=0 is Start, Desired=1 is Stop. Generic action query is Stop.
           IF #Desired = 0 THEN
               IF #Unit.Mode = 1 OR #Unit.ModePending THEN
                   "FRK_ReleaseReason"(Report := #Report,
                                       Description := WSTRING#'std.error.unsupportedModeRequest',
                                       Reason := 2002,
                                       Path := STRING_TO_WSTRING(#Status.Name),
                                       Kind := 0);
               END_IF;
               IF #Core.Exec <> 0 OR #Unit.RunReq OR #Unit.Clearing OR #Unit.FaultLatched THEN
                   "FRK_ReleaseReason"(Report := #Report,
                                       Description := WSTRING#'std.error.hmiRequestRejected',
                                       Reason := 2011,
                                       Path := STRING_TO_WSTRING(#Status.Name),
                                       Kind := 4);
               END_IF;
               IF #Unit.AlarmBlocking THEN
                   "FRK_ReleaseReason"(Report := #Report,
                                       Description := WSTRING#'std.release.manualReset',
                                       Reason := 0,
                                       Path := STRING_TO_WSTRING(#Status.Name),
                                       Kind := 2);
               END_IF;
               IF #Unit.ConfigBlocked THEN
                   "FRK_ReleaseReason"(Report := #Report,
                                       Description := WSTRING#'std.release.configRestoreUnacknowledged',
                                       Reason := 2040,
                                       Path := STRING_TO_WSTRING(#Status.Name),
                                       Kind := 2);
               END_IF;
               IF NOT #Unit.Permit THEN
                   "FRK_ReleaseReason"(Report := #Report,
                                       Description := #Unit.PermitDiag.Description,
                                       Reason := #Unit.PermitDiag.ReasonCode,
                                       Path := #Unit.PermitDiag.SourcePath,
                                       Kind := 3);
               END_IF;
           END_IF;
       4:
           IF #Unit.ModePending THEN
               "FRK_ReleaseReason"(Report := #Report,
                                   Description := WSTRING#'std.release.modeChangeAlreadyPending',
                                   Reason := 2011,
                                   Path := STRING_TO_WSTRING(#Status.Name),
                                   Kind := 0);
           END_IF;
           IF #Core.Exec = 1 AND #Unit.Mode <> 1 THEN
               IF #Policy[#Unit.Mode].Shield = 2 THEN
                   "FRK_ReleaseReason"(Report := #Report,
                                       Description := WSTRING#'std.release.modeSwitchBlockedWhileRunning',
                                       Reason := 2002,
                                       Path := STRING_TO_WSTRING(#Status.Name),
                                       Kind := 0);
               END_IF;
           END_IF;
           IF #Desired <> -1 THEN
               IF #Desired < 0 OR #Desired >= 7 THEN
                   "FRK_ReleaseReason"(Report := #Report,
                                       Description := WSTRING#'std.error.unsupportedModeRequest',
                                       Reason := 2008,
                                       Path := STRING_TO_WSTRING(#Status.Name),
                                       Kind := 0);
               ELSIF NOT #Supported[#Desired] THEN
                   "FRK_ReleaseReason"(Report := #Report,
                                       Description := WSTRING#'std.error.unsupportedModeRequest',
                                       Reason := 2008,
                                       Path := STRING_TO_WSTRING(#Status.Name),
                                       Kind := 0);
               END_IF;
           END_IF;
       7:
           // The complete alarm model is separate; this gate owns the current latch.
           IF NOT #Unit.FaultLatched AND NOT #Unit.AlarmBlocking AND #Core.Exec = 0 AND NOT #Unit.Clearing AND NOT #Unit.ModePending AND NOT #Unit.FollowStart THEN
               IF "FRK_DescendantsReady"(OwnerIndex := #Core.RegIndex) THEN
                   "FRK_ReleaseReason"(Report := #Report,
                                       Description := WSTRING#'std.release.noBlockingAlarm',
                                       Reason := 2011,
                                       Path := STRING_TO_WSTRING(#Status.Name),
                                       Kind := 4);
               END_IF;
           END_IF;
       2:
           "FRK_ManualCommon"(Core := #Core,
                              Unit := #Unit,
                              Status := #Status,
                              Report := #Report);
       ELSE
           RETURN;
   END_CASE;
END_FUNCTION

FUNCTION "FRK_UnitRunStart" : Void   // FC83, SCL
{ S7_Optimized_Access := 'TRUE' }
VERSION : 0.1
// stored: AutoNumber true, IsIECCheckEnabled false, SetENOAutomatically false, UDAEnableTagReadback false
   VAR_INPUT
      Timeout : Time;
      Label : String;
   END_VAR
   VAR_IN_OUT
      Core : "FRK_Core";
      Status : "ST_ModuleStatus";
   END_VAR
BEGIN

   "FRK_Start"(Core := #Core,
               Status := #Status,
               Supported := TRUE,
               Timeout := #Timeout,
               Label := #Label);
   // A continuous run ends at Stop. Bounded commands/steps own progress timeouts.
   #Core.TimeoutMs := 0;
END_FUNCTION

FUNCTION "FRK_UnitSetLocalCarrier" : Void   // FC70, SCL
{ S7_Optimized_Access := 'TRUE' }
VERSION : 0.1
// stored: AutoNumber true, IsIECCheckEnabled false, SetENOAutomatically false, UDAEnableTagReadback false
   VAR_INPUT
      Index : DInt;
   END_VAR
   VAR_IN_OUT
      Unit : "FRK_Unit";
   END_VAR
BEGIN

   #Unit.CarrierIndex := 0;
   IF #Index < 1 OR #Index > 32 THEN
       RETURN;
   END_IF;
   "FRK_Carriers".Slots[#Index].Enabled := TRUE;
   "FRK_Carriers".Slots[#Index].Kind := 2;
   #Unit.CarrierIndex := #Index;
END_FUNCTION

FUNCTION "FRK_UnitSetPermit" : Void   // FC76, SCL
{ S7_Optimized_Access := 'TRUE' }
VERSION : 0.1
// stored: AutoNumber true, IsIECCheckEnabled false, SetENOAutomatically false, UDAEnableTagReadback false
   VAR_INPUT
      Ok : Bool;
      Diag : "ST_Diagnostic";
   END_VAR
   VAR_IN_OUT
      Unit : "FRK_Unit";
   END_VAR
BEGIN

   #Unit.Permit := #Ok;
   #Unit.PermitDiag := #Diag;
END_FUNCTION

FUNCTION "F_AccessBenchProvision" : Void   // FC176, SCL
{ S7_Optimized_Access := 'TRUE' }
VERSION : 0.1
// stored: AutoNumber true, IsIECCheckEnabled false, SetENOAutomatically false, UDAEnableTagReadback false
BEGIN

   "FRK_LocalUsers".Count := 2;
   "FRK_LocalUsers".Rows[1].User := 'operator';
   "FRK_LocalUsers".Rows[1].Level := 1;
   "FRK_LocalUsers".Rows[1].Salt[0] := BYTE#16#75;
   "FRK_LocalUsers".Rows[1].Salt[1] := BYTE#16#C6;
   "FRK_LocalUsers".Rows[1].Salt[2] := BYTE#16#08;
   "FRK_LocalUsers".Rows[1].Salt[3] := BYTE#16#35;
   "FRK_LocalUsers".Rows[1].Salt[4] := BYTE#16#0C;
   "FRK_LocalUsers".Rows[1].Salt[5] := BYTE#16#C0;
   "FRK_LocalUsers".Rows[1].Salt[6] := BYTE#16#0E;
   "FRK_LocalUsers".Rows[1].Salt[7] := BYTE#16#9A;
   "FRK_LocalUsers".Rows[1].Salt[8] := BYTE#16#16;
   "FRK_LocalUsers".Rows[1].Salt[9] := BYTE#16#1E;
   "FRK_LocalUsers".Rows[1].Salt[10] := BYTE#16#4A;
   "FRK_LocalUsers".Rows[1].Salt[11] := BYTE#16#85;
   "FRK_LocalUsers".Rows[1].Salt[12] := BYTE#16#D4;
   "FRK_LocalUsers".Rows[1].Salt[13] := BYTE#16#41;
   "FRK_LocalUsers".Rows[1].Salt[14] := BYTE#16#E9;
   "FRK_LocalUsers".Rows[1].Salt[15] := BYTE#16#3E;
   "FRK_LocalUsers".Rows[1].PinHash[0] := BYTE#16#D1;
   "FRK_LocalUsers".Rows[1].PinHash[1] := BYTE#16#62;
   "FRK_LocalUsers".Rows[1].PinHash[2] := BYTE#16#D8;
   "FRK_LocalUsers".Rows[1].PinHash[3] := BYTE#16#FC;
   "FRK_LocalUsers".Rows[1].PinHash[4] := BYTE#16#F2;
   "FRK_LocalUsers".Rows[1].PinHash[5] := BYTE#16#CE;
   "FRK_LocalUsers".Rows[1].PinHash[6] := BYTE#16#BA;
   "FRK_LocalUsers".Rows[1].PinHash[7] := BYTE#16#54;
   "FRK_LocalUsers".Rows[1].PinHash[8] := BYTE#16#13;
   "FRK_LocalUsers".Rows[1].PinHash[9] := BYTE#16#AF;
   "FRK_LocalUsers".Rows[1].PinHash[10] := BYTE#16#4D;
   "FRK_LocalUsers".Rows[1].PinHash[11] := BYTE#16#AC;
   "FRK_LocalUsers".Rows[1].PinHash[12] := BYTE#16#ED;
   "FRK_LocalUsers".Rows[1].PinHash[13] := BYTE#16#2A;
   "FRK_LocalUsers".Rows[1].PinHash[14] := BYTE#16#DF;
   "FRK_LocalUsers".Rows[1].PinHash[15] := BYTE#16#A6;
   "FRK_LocalUsers".Rows[1].PinHash[16] := BYTE#16#0D;
   "FRK_LocalUsers".Rows[1].PinHash[17] := BYTE#16#EE;
   "FRK_LocalUsers".Rows[1].PinHash[18] := BYTE#16#80;
   "FRK_LocalUsers".Rows[1].PinHash[19] := BYTE#16#98;
   "FRK_LocalUsers".Rows[1].PinHash[20] := BYTE#16#6C;
   "FRK_LocalUsers".Rows[1].PinHash[21] := BYTE#16#2F;
   "FRK_LocalUsers".Rows[1].PinHash[22] := BYTE#16#92;
   "FRK_LocalUsers".Rows[1].PinHash[23] := BYTE#16#84;
   "FRK_LocalUsers".Rows[1].PinHash[24] := BYTE#16#2D;
   "FRK_LocalUsers".Rows[1].PinHash[25] := BYTE#16#66;
   "FRK_LocalUsers".Rows[1].PinHash[26] := BYTE#16#38;
   "FRK_LocalUsers".Rows[1].PinHash[27] := BYTE#16#1E;
   "FRK_LocalUsers".Rows[1].PinHash[28] := BYTE#16#5B;
   "FRK_LocalUsers".Rows[1].PinHash[29] := BYTE#16#33;
   "FRK_LocalUsers".Rows[1].PinHash[30] := BYTE#16#2B;
   "FRK_LocalUsers".Rows[1].PinHash[31] := BYTE#16#94;
   "FRK_LocalUsers".Rows[2].User := 'admin';
   "FRK_LocalUsers".Rows[2].Level := 4;
   "FRK_LocalUsers".Rows[2].Salt[0] := BYTE#16#2C;
   "FRK_LocalUsers".Rows[2].Salt[1] := BYTE#16#11;
   "FRK_LocalUsers".Rows[2].Salt[2] := BYTE#16#7A;
   "FRK_LocalUsers".Rows[2].Salt[3] := BYTE#16#95;
   "FRK_LocalUsers".Rows[2].Salt[4] := BYTE#16#98;
   "FRK_LocalUsers".Rows[2].Salt[5] := BYTE#16#C1;
   "FRK_LocalUsers".Rows[2].Salt[6] := BYTE#16#2A;
   "FRK_LocalUsers".Rows[2].Salt[7] := BYTE#16#CF;
   "FRK_LocalUsers".Rows[2].Salt[8] := BYTE#16#BC;
   "FRK_LocalUsers".Rows[2].Salt[9] := BYTE#16#6E;
   "FRK_LocalUsers".Rows[2].Salt[10] := BYTE#16#06;
   "FRK_LocalUsers".Rows[2].Salt[11] := BYTE#16#4E;
   "FRK_LocalUsers".Rows[2].Salt[12] := BYTE#16#17;
   "FRK_LocalUsers".Rows[2].Salt[13] := BYTE#16#E6;
   "FRK_LocalUsers".Rows[2].Salt[14] := BYTE#16#5E;
   "FRK_LocalUsers".Rows[2].Salt[15] := BYTE#16#43;
   "FRK_LocalUsers".Rows[2].PinHash[0] := BYTE#16#FD;
   "FRK_LocalUsers".Rows[2].PinHash[1] := BYTE#16#4F;
   "FRK_LocalUsers".Rows[2].PinHash[2] := BYTE#16#56;
   "FRK_LocalUsers".Rows[2].PinHash[3] := BYTE#16#ED;
   "FRK_LocalUsers".Rows[2].PinHash[4] := BYTE#16#D8;
   "FRK_LocalUsers".Rows[2].PinHash[5] := BYTE#16#A6;
   "FRK_LocalUsers".Rows[2].PinHash[6] := BYTE#16#58;
   "FRK_LocalUsers".Rows[2].PinHash[7] := BYTE#16#AA;
   "FRK_LocalUsers".Rows[2].PinHash[8] := BYTE#16#B6;
   "FRK_LocalUsers".Rows[2].PinHash[9] := BYTE#16#AF;
   "FRK_LocalUsers".Rows[2].PinHash[10] := BYTE#16#D9;
   "FRK_LocalUsers".Rows[2].PinHash[11] := BYTE#16#91;
   "FRK_LocalUsers".Rows[2].PinHash[12] := BYTE#16#87;
   "FRK_LocalUsers".Rows[2].PinHash[13] := BYTE#16#D5;
   "FRK_LocalUsers".Rows[2].PinHash[14] := BYTE#16#18;
   "FRK_LocalUsers".Rows[2].PinHash[15] := BYTE#16#EF;
   "FRK_LocalUsers".Rows[2].PinHash[16] := BYTE#16#A5;
   "FRK_LocalUsers".Rows[2].PinHash[17] := BYTE#16#79;
   "FRK_LocalUsers".Rows[2].PinHash[18] := BYTE#16#BA;
   "FRK_LocalUsers".Rows[2].PinHash[19] := BYTE#16#82;
   "FRK_LocalUsers".Rows[2].PinHash[20] := BYTE#16#87;
   "FRK_LocalUsers".Rows[2].PinHash[21] := BYTE#16#7E;
   "FRK_LocalUsers".Rows[2].PinHash[22] := BYTE#16#F4;
   "FRK_LocalUsers".Rows[2].PinHash[23] := BYTE#16#C3;
   "FRK_LocalUsers".Rows[2].PinHash[24] := BYTE#16#47;
   "FRK_LocalUsers".Rows[2].PinHash[25] := BYTE#16#A5;
   "FRK_LocalUsers".Rows[2].PinHash[26] := BYTE#16#95;
   "FRK_LocalUsers".Rows[2].PinHash[27] := BYTE#16#2E;
   "FRK_LocalUsers".Rows[2].PinHash[28] := BYTE#16#AB;
   "FRK_LocalUsers".Rows[2].PinHash[29] := BYTE#16#60;
   "FRK_LocalUsers".Rows[2].PinHash[30] := BYTE#16#10;
   "FRK_LocalUsers".Rows[2].PinHash[31] := BYTE#16#C4;

   "GDB_AccessPersistTest".ProvisionCount := "GDB_AccessPersistTest".ProvisionCount + 1;
END_FUNCTION

FUNCTION "F_AccessPersistenceBench" : Void   // FC174, SCL
{ S7_Optimized_Access := 'TRUE' }
VERSION : 0.1
// Deliberate engineering-only stimuli. Never generated into a station.
// stored: AutoNumber true, IsIECCheckEnabled false, SetENOAutomatically false, UDAEnableTagReadback false
   VAR_INPUT
      Startup : Bool;
   END_VAR
   VAR_TEMP
      Index : Int;
      Accepted : Bool;
      Crc : DWord;
      Vector : String[9];
   END_VAR
BEGIN

   IF #Startup THEN
       "GDB_AccessPersistTest".StartupCount := "GDB_AccessPersistTest".StartupCount + 1;
       #Vector := '123456789';
       #Crc := DWORD#16#FFFFFFFF;
       FOR #Index := 1 TO 9 DO
           #Crc := "FRK_CrcByte"(Previous := #Crc, Value := CHAR_TO_BYTE(#Vector[#Index]));
       END_FOR;
       "GDB_AccessPersistTest".CrcWitness := NOT #Crc;
   END_IF;
   IF "GDB_AccessPersistTest".RotateOnLogin AND "StationA".Access.LoginBusy THEN
       "GDB_AccessPersistTest".Operation := 1;
       "GDB_AccessPersistTest".RotateOnLogin := FALSE;
   END_IF;
   IF "GDB_AccessPersistTest".Operation <> 0 THEN
       "GDB_AccessPersistTest".Applied := FALSE;
       "GDB_AccessPersistTest".PolicySlot := 0;
       FOR #Index := 1 TO 2 DO
           IF "FRK_AccessPolicies".Rows[#Index].Scope = "GDB_AccessPersistTest".Root THEN
               "GDB_AccessPersistTest".PolicySlot := #Index;
           END_IF;
       END_FOR;
       CASE "GDB_AccessPersistTest".Operation OF
           1: // Real trusted registration: edit the operator role, preserving its salted hash.
               "GDB_AccessPersistTest".Record := "FRK_LocalUsers".Rows[1];
               "GDB_AccessPersistTest".Record.Level := "GDB_AccessPersistTest".Value;
               "GDB_AccessPersistTest".Applied := "FRK_AccessRegisterHash"(Record := "GDB_AccessPersistTest".Record);
           2:
               "FRK_LocalUsers".SchemaVersion := DINT_TO_UINT("GDB_AccessPersistTest".Value);
               "GDB_AccessPersistTest".Applied := TRUE;
           3:
               "FRK_LocalUsers".Count := "GDB_AccessPersistTest".Value;
               "GDB_AccessPersistTest".Applied := TRUE;
           4:
               "FRK_LocalUsers".Rows[1].Level := "GDB_AccessPersistTest".Value;
               "GDB_AccessPersistTest".Applied := TRUE;
           5:
               "FRK_LocalUsers".Rows[1].User := "FRK_LocalUsers".Rows[2].User;
               "GDB_AccessPersistTest".Applied := TRUE;
           6:
               "FRK_LocalUsers".Rows[1].PinHash[31] := "FRK_LocalUsers".Rows[1].PinHash[31] XOR BYTE#1;
               "GDB_AccessPersistTest".Applied := TRUE;
           7: "F_AccessBenchProvision"();
               "GDB_AccessPersistTest".Applied := "FRK_AccessUsersCommit"();
           8:
               "FRK_LocalUsers".SchemaVersion := 0;
               "FRK_LocalUsers".Generation := 0;
               "FRK_LocalUsers".Checksum := DWORD#0;
               "GDB_AccessPersistTest".Applied := TRUE;
           10, 11, 12, 13:
               IF "GDB_AccessPersistTest".PolicySlot > 0 THEN
                   CASE "GDB_AccessPersistTest".Operation OF
                       10:
                           "FRK_AccessPolicies".Rows["GDB_AccessPersistTest".PolicySlot].SchemaVersion := DINT_TO_UINT("GDB_AccessPersistTest".Value);
                       11:
                           "FRK_AccessPolicies".Rows["GDB_AccessPersistTest".PolicySlot].Policy.Required["GDB_AccessPersistTest".Gate] := "GDB_AccessPersistTest".Value;
                       13:
                           "FRK_AccessPolicies".Rows["GDB_AccessPersistTest".PolicySlot].SchemaVersion := 0;
                           "FRK_AccessPolicies".Rows["GDB_AccessPersistTest".PolicySlot].Generation := 0;
                           "FRK_AccessPolicies".Rows["GDB_AccessPersistTest".PolicySlot].Checksum := DWORD#0;
                       12:
                           "FRK_AccessPolicies".Rows["GDB_AccessPersistTest".PolicySlot].Checksum := "FRK_AccessPolicies".Rows["GDB_AccessPersistTest".PolicySlot].Checksum XOR DWORD#1;
                   END_CASE;
                   "GDB_AccessPersistTest".Applied := TRUE;
               END_IF;
       END_CASE;
       "GDB_AccessPersistTest".Operation := 0;
   END_IF;
   "GDB_AccessPersistTest".UsersReady := "FRK_AccessStorage".UsersReady;
   "GDB_AccessPersistTest".UsersLost := "FRK_AccessStorage".UsersLost;
   "GDB_AccessPersistTest".UserGeneration := "FRK_LocalUsers".Generation;
END_FUNCTION

FUNCTION "F_AlarmPersistenceBench" : Void   // FC175, SCL
{ S7_Optimized_Access := 'TRUE' }
VERSION : 0.1
// stored: AutoNumber true, IsIECCheckEnabled false, SetENOAutomatically false, UDAEnableTagReadback false
   VAR_TEMP
      Slot : Int;
   END_VAR
BEGIN

   #Slot := "FRK_AlarmHistoryIndex"(Scope := "GDB_AlarmPersistTest".Scope);
   "GDB_AlarmPersistTest".Slot := #Slot;
   IF #Slot < 1 THEN
       RETURN;
   END_IF;
   "GDB_AlarmPersistTest".Generation := "FRK_AlarmHistory".Rows[#Slot].Generation;
   "GDB_AlarmPersistTest".Checksum := "FRK_AlarmHistory".Rows[#Slot].Checksum;
   "GDB_AlarmPersistTest".Used := "FRK_AlarmHistory".Rows[#Slot].RingUsed;
   "GDB_AlarmPersistTest".Applied := "GDB_AlarmPersistTest".Operation <> 0;
   CASE "GDB_AlarmPersistTest".Operation OF
       1, 2:
           IF "GDB_AlarmPersistTest".Scope = 'StationA' THEN
               IF "GDB_AlarmPersistTest".Operation = 1 THEN
                   "FRK_AlarmMessage"(Reason := "GDB_AlarmPersistTest".Reason,
                                      Description := "GDB_AlarmPersistTest".Text,
                                      SourcePath := WSTRING#'StationA',
                                      AlarmLog := "StationA".AlarmLog);
               ELSE
                   "FRK_AlarmBegin"(Startup := TRUE,
                                    AlarmLog := "StationA".AlarmLog);
               END_IF;
           END_IF;
           IF "GDB_AlarmPersistTest".Scope = 'StationA.Satellite' THEN
               IF "GDB_AlarmPersistTest".Operation = 1 THEN
                   "FRK_AlarmMessage"(Reason := "GDB_AlarmPersistTest".Reason,
                                      Description := "GDB_AlarmPersistTest".Text,
                                      SourcePath := WSTRING#'StationA.Satellite',
                                      AlarmLog := "StationA".Satellite.AlarmLog);
               ELSE
                   "FRK_AlarmBegin"(Startup := TRUE,
                                    AlarmLog := "StationA".Satellite.AlarmLog);
               END_IF;
           END_IF;
           IF "GDB_AlarmPersistTest".Scope = 'StationA.Satellite.Inner' THEN
               IF "GDB_AlarmPersistTest".Operation = 1 THEN
                   "FRK_AlarmMessage"(Reason := "GDB_AlarmPersistTest".Reason,
                                      Description := "GDB_AlarmPersistTest".Text,
                                      SourcePath := WSTRING#'StationA.Satellite.Inner',
                                      AlarmLog := "StationA".Satellite.Inner.AlarmLog);
               ELSE
                   "FRK_AlarmBegin"(Startup := TRUE,
                                    AlarmLog := "StationA".Satellite.Inner.AlarmLog);
               END_IF;
           END_IF;
           IF "GDB_AlarmPersistTest".Scope = 'StationB' THEN
               IF "GDB_AlarmPersistTest".Operation = 1 THEN
                   "FRK_AlarmMessage"(Reason := "GDB_AlarmPersistTest".Reason,
                                      Description := "GDB_AlarmPersistTest".Text,
                                      SourcePath := WSTRING#'StationB',
                                      AlarmLog := "StationB".AlarmLog);
               ELSE
                   "FRK_AlarmBegin"(Startup := TRUE,
                                    AlarmLog := "StationB".AlarmLog);
               END_IF;
           END_IF;
           IF "GDB_AlarmPersistTest".Scope = 'StationB.Satellite' THEN
               IF "GDB_AlarmPersistTest".Operation = 1 THEN
                   "FRK_AlarmMessage"(Reason := "GDB_AlarmPersistTest".Reason,
                                      Description := "GDB_AlarmPersistTest".Text,
                                      SourcePath := WSTRING#'StationB.Satellite',
                                      AlarmLog := "StationB".Satellite.AlarmLog);
               ELSE
                   "FRK_AlarmBegin"(Startup := TRUE,
                                    AlarmLog := "StationB".Satellite.AlarmLog);
               END_IF;
           END_IF;
           IF "GDB_AlarmPersistTest".Scope = 'StationB.Satellite.Inner' THEN
               IF "GDB_AlarmPersistTest".Operation = 1 THEN
                   "FRK_AlarmMessage"(Reason := "GDB_AlarmPersistTest".Reason,
                                      Description := "GDB_AlarmPersistTest".Text,
                                      SourcePath := WSTRING#'StationB.Satellite.Inner',
                                      AlarmLog := "StationB".Satellite.Inner.AlarmLog);
               ELSE
                   "FRK_AlarmBegin"(Startup := TRUE,
                                    AlarmLog := "StationB".Satellite.Inner.AlarmLog);
               END_IF;
           END_IF;
       10:
           "FRK_AlarmHistory".Rows[#Slot].SchemaVersion := 2;
       11:
           "FRK_AlarmHistory".Rows[#Slot].RingHead := 65;
       12:
           "FRK_AlarmHistory".Rows[#Slot].Checksum := "FRK_AlarmHistory".Rows[#Slot].Checksum XOR DWORD#1;
       13:
           "FRK_AlarmHistory".Rows[#Slot].Scope := 'foreign';
       14:
           "FRK_AlarmHistory".Rows[#Slot].Ring[1].Description := WSTRING#'corrupted';
       15:
           "FRK_AlarmHistory".Rows[#Slot].Ring[1].Duration := T#-1ms;
       16:
           "FRK_AlarmHistory".Rows[#Slot].SchemaVersion := 0;
           "FRK_AlarmHistory".Rows[#Slot].Generation := 0;
           "FRK_AlarmHistory".Rows[#Slot].Scope := '';
           "FRK_AlarmHistory".Rows[#Slot].Checksum := DWORD#0;
       17:
           "FRK_AlarmHistory".Rows[#Slot].RingUsed := -1;
   END_CASE;
   "GDB_AlarmPersistTest".Operation := 0;
END_FUNCTION

FUNCTION "F_ConfigBenchObserve" : Void   // FC178, SCL
{ S7_Optimized_Access := 'TRUE' }
VERSION : 0.1
// stored: AutoNumber true, IsIECCheckEnabled false, SetENOAutomatically false, UDAEnableTagReadback false
   VAR_INPUT
      Startup : Bool;
   END_VAR
BEGIN

   "GDB_StateAlarmTest".NativeFaultSlot := "StationA".Cell.Gate.Core.FaultSlot;
   "GDB_RoutingTest".ManExecute := "StationA".Cell.Gate.Execute;
   "GDB_RoutingTest".ManStarts := "StationA".Cell.Gate.Device.StartCount;
   "GDB_UnitTest".Scans := "GDB_UnitTest".Scans + 1;
   "GDB_UnitTest".ChildExecute := "StationA".Cell.Clamp.Execute;
   "GDB_UnitTest".ChildState := "StationA".Cell.Clamp.Core.Exec;
   "GDB_UnitTest".CarrierWrites := "FRK_Carriers".Slots[1].Writes;
   "GDB_UnitTest".CarrierSerial := "FRK_Carriers".Slots[1].Serial;
   "GDB_UnitTest".WrittenUid := "FRK_Carriers".Slots[1].Written.Uid;
   "GDB_UnitTest".WrittenVerdict := "FRK_Carriers".Slots[1].Written.Result.Verdict;
   IF "StationA".AlarmLog.RingHead > 0 AND "StationA".AlarmLog.RingHead <= 64 THEN
       "GDB_UnitTest".LastEvent := "StationA".AlarmLog.Ring["StationA".AlarmLog.RingHead].ReasonCode;
   END_IF;
   "GDB_UnitTest".SecretCleared := "StationA".HmiRequest.Secret = '';
   "GDB_UnitTest".SnapshotSecretCleared := "StationA".Unit.Request.Secret = '';
   IF "StationA".Access.LoginBusy AND ("GDB_AccessTest".CancelOnLogin OR "GDB_AccessTest".SupersedeOnLogin) THEN
       "GDB_AccessTest".InterruptedBusy := TRUE;
       IF "GDB_AccessTest".CancelOnLogin THEN
           "GDB_AccessTest".InterruptRequest.Kind := 2;
           "FRK_UnitOperation"(Core := "StationA".Core,
                               Unit := "StationA".Unit,
                               Status := "StationA".Status,
                               Policy := "StationA".ModePolicy,
                               Access := "StationA".Access,
                               Supported := "StationA".SupportedModesPublished,
                               Request := "GDB_AccessTest".InterruptRequest,
                               Response := "FRK_UnitScratch".Response,
                               Trusted := FALSE);
       ELSE
           "GDB_AccessTest".SupersededSequence := "FRK_AccessNext"(Previous := "StationA".Access.LoginSequence);
           "FRK_AccessLogin"(Access := "StationA".Access,
                             User := 'unknown',
                             Secret := 'wrong',
                             Sequence := "GDB_AccessTest".SupersededSequence);
       END_IF;
       "GDB_AccessTest".CancelOnLogin := FALSE;
       "GDB_AccessTest".SupersedeOnLogin := FALSE;
   END_IF;
   "F_ConfigSetBench"();
   "F_AccessPersistenceBench"(Startup := #Startup);
   "F_AlarmPersistenceBench"();
END_FUNCTION

FUNCTION "F_ConfigBenchPrepare" : Void   // FC177, SCL
{ S7_Optimized_Access := 'TRUE' }
VERSION : 0.1
// stored: AutoNumber true, IsIECCheckEnabled false, SetENOAutomatically false, UDAEnableTagReadback false
   VAR_INPUT
      Startup : Bool;
   END_VAR
   VAR_TEMP
      StartupStamp : DTL;
      ResultCode : Int;
      SlotIndex : Int;
      Taken : Int;
      Accepted : Bool;
   END_VAR
BEGIN

